// TIA Portal V21 export
// export: Created 2026-08-21T20:18:51.8937952Z, ExportSetting None, DisplayName Totally Integrated Automation Portal, DisplayVersion V21, DisplayName STEP 7 Professional, DisplayVersion V21, DisplayName STEP 7 Safety, DisplayVersion V21, DisplayName Tech WebApplication, DisplayVersion V21, DisplayName WinCC Basic/Comfort/Advanced, DisplayVersion V21, DisplayName WinCC Professional, DisplayVersion V21, DisplayName WinCC Unified, DisplayVersion V21
DATA_BLOCK "ConfigurationParameters_DB"   // DB32
AUTHOR : Siemens AG
FAMILY : ServiceControl
VERSION : 1.0
// stored: InstanceOfName ConfigurationParameters, InstanceOfType FB
"ConfigurationParameters"
   // VAR
   //    MTPAnalog { S7_SetPoint := 'True'} : Array[0..0] of "UDT_MTP_AnaServParam";
   //    MTPDigital { S7_SetPoint := 'True'} : Array[0..0] of "UDT_MTP_DIntServParam";
   //    MTPBinary { S7_SetPoint := 'True'} : Array[0..1] of "UDT_MTP_BinServParam";
   //    MTPString { S7_SetPoint := 'True'} : Array[0..0] of "UDT_MTP_StringServParam";
   // END_VAR
BEGIN
   MTPBinary[0].VExt := True;
   MTPBinary[0].VOp := True;
   MTPBinary[0].VInt := True;
   MTPBinary[0].VReq := True;
   MTPBinary[0].VOut := True;
   MTPBinary[0].VState0 := 'Other PEA not co';
   MTPBinary[0].VState1 := 'Other PEA connec';
END_DATA_BLOCK
